Staubli VAL3: Lab2A_L1.dtx


